(* IEC 61131-3 sources: plc_generation_empirical_study/datasets/packages/internal_v0_1/qualification_only/C03_E01_forward_reverse_interlock, 1 file *)

(* ---- reference.st ---- *)
FUNCTION_BLOCK C03_E01_forward_reverse_interlock
VAR_INPUT
    ForwardRequest : BOOL;
    ReverseRequest : BOOL;
    Permit : BOOL;
END_VAR
VAR_OUTPUT
    Forward : BOOL;
    Reverse : BOOL;
END_VAR

Forward := Permit AND ForwardRequest AND (NOT ReverseRequest);
Reverse := Permit AND ReverseRequest AND (NOT ForwardRequest);

END_FUNCTION_BLOCK
